(* IEC 61131-3 sources: llm-plc-st-eval/data/processed_definitivo/gemini-3.1-pro-preview/B7/zero_shot, 3 files *)

(* ---- ejec_1.st ---- *)
FUNCTION SelBomba : BOOL
VAR_INPUT
    modoAuto : BOOL;  (* TRUE = Modo Automático, FALSE = Modo Manual *)
    btnManual : BOOL; (* Comando de encendido en modo manual *)
    nivelBajo : BOOL; (* Condición de encendido en modo automático *)
END_VAR

(*
   Al ser una lógica puramente combinacional sin memoria entre ciclos,
   el tipo de POU más adecuado es una FUNCTION. El resultado se
   devuelve en el propio nombre de la función.
*)
SelBomba := (modoAuto AND nivelBajo) OR (NOT modoAuto AND btnManual);

END_FUNCTION

(* ---- ejec_2.st ---- *)
FUNCTION SelBomba : BOOL
VAR_INPUT
    modoAuto : BOOL;  // TRUE = Modo Automático, FALSE = Modo Manual
    btnManual : BOOL; // Comando directo de la bomba en modo manual
    nivelBajo : BOOL; // Condición para encender la bomba en modo automático
END_VAR

(*
   Al ser una lógica puramente combinacional sin memoria entre ciclos,
   una FUNCTION es la POU más adecuada. El estado de la bomba se
   asigna directamente al valor de retorno de la función (SelBomba).
*)

SelBomba := (modoAuto AND nivelBajo) OR (NOT modoAuto AND btnManual);

END_FUNCTION

(* ---- ejec_3.st ---- *)
FUNCTION SelBomba : BOOL
VAR_INPUT
    modoAuto : BOOL;  // TRUE = Modo Automático, FALSE = Modo Manual
    btnManual : BOOL; // Comando de encendido en modo manual
    nivelBajo : BOOL; // Condición de encendido en modo automático
END_VAR

(*
   Al no requerir memoria entre ciclos (lógica puramente combinacional),
   una FUNCTION es la unidad de organización de programa (POU) más adecuada.
*)

IF modoAuto THEN
    // En modo automático, el estado depende de la señal de nivel bajo
    SelBomba := nivelBajo;
ELSE
    // En modo manual, el estado obedece directamente al botón
    SelBomba := btnManual;
END_IF;

// Nota: También se puede expresar como:
// SelBomba := (modoAuto AND nivelBajo) OR (NOT modoAuto AND btnManual);

END_FUNCTION
